(* IEC 61131-3 sources: programs/VI-54/VI-54_20171205/VI-54_20171205/Stations/PLC_VI54/VI-54_171014/Class/_DriveAxisBase (part 2) *)

  //Error of Axis gets only shown, if Axis is Online
  if bOnlineFinished then
    AxError := GetAxError();
  else
    AxError := 0;
  end_if;

  output := AxError;

END_FUNCTION

FUNCTION _DriveAxisBase::LoadDrivePara
  VAR
    pTabAdress : ^DINT;
    TabLength   : DINT;
  END_VAR

  // load the parameter data to the para objects
  case DriveInitType of

    _SDDSTDTABLE :

     pTabAdress := GetTabAdress(TabType:= 0, bdSettings.bSendMPara, #TabLength);
     SetListToParObj(pData:= (pTabAdress)$^DINT, udLen:=TabLength$UDINT);

    _SDDL2TABLE :
    // load the data of the table
      pTabAdress := GetTabAdress(TabType:= 1, bdSettings.bSendMPara, #TabLength);
      SetListToParObj(pData:= (pTabAdress)$^DINT, udLen:=TabLength$UDINT);

    _SDDRAMEX,
    _SDDFILE :
      pSDDData$^void := DriveAxisSet.GetMemPtr();
      if pSDDData <> NIL then
        // load the data of the memory
        SetListToParObj(pData:= (pSDDData$DINT + pSDDData^.AxOffset)$^DINT, udLen:=pSDDData^.AxLength);
      end_if;

  end_case;

END_FUNCTION

FUNCTION _DriveAxisBase::SetListToParObj
	VAR_INPUT
		pData 	: ^DINT;
		udLen 	: UDINT;
	END_VAR
	VAR_OUTPUT
		retcode 	: BOOL;
	END_VAR
  VAR
    pHlp          : ^DINT;
    x             : UDINT;
    pThisNewInst  : ^void;
    usParaNr      : USINT;
    ParaValue     : DINT;
    UserPara      : CmdStruct;
    UserResult    : Results;
  END_VAR

  retcode := FALSE;

  //hier konnte es zu einem Problem kommen kann wenn pThisNewInst nicht init war.
  pThisNewInst := NIL; //BleErn 19.08.2010 11:27

  if (bdSettings.bAxSetPara = FALSE) | (pData = NIL) then
    return;
  end_if;

  x := 0;
  pHlp := pData;

  while x < udLen do

    usParaNr := pHlp^$USINT;
    pHlp += sizeof(USINT);
    x += sizeof(USINT);

    if usParaNr <= MAX_MOTOR_PARA then
      pThisNewInst$DINT := AxSetPara[IDX_MOTOR_PARA];
    elsif usParaNr <= MAX_DRIVE_PARA then
      pThisNewInst$DINT := AxSetPara[IDX_DRIVE_PARA];
    elsif usParaNr <= MAX_CURRENT_PARA then
      pThisNewInst$DINT := AxSetPara[IDX_CURRENT_PARA];
    elsif usParaNr <= MAX_VEL_PARA then
      pThisNewInst$DINT := AxSetPara[IDX_VEL_PARA];
    elsif usParaNr <= MAX_POS_PARA then
      pThisNewInst$DINT := AxSetPara[IDX_POS_PARA];
    elsif usParaNr <= MAX_FD_PARA then
      pThisNewInst$DINT := AxSetPara[IDX_FD_PARA];
    elsif usParaNr <= MAX_APPLI_PARA then
      pThisNewInst$DINT := AxSetPara[IDX_APPLI_PARA];
    elsif usParaNr <= MAX_ERRORHANDLING then
      pThisNewInst$DINT := AxSetPara[IDX_ERRORHANDLING];
    end_if;

    ParaValue := pHlp^$DINT;
    if pThisNewInst <> NIL then
      UserPara.uiCmd := SDD_REFRESH_SETPARA;
      UserPara.aPara[0] := to_dint(usParaNr);
      UserPara.aPara[1] := ParaValue;
      pThisNewInst$^VirtualBase^.NewInst(#UserPara, #UserResult);
    end_if;

    pHlp += sizeof(UDINT);
    x += sizeof(UDINT);

  end_while;

END_FUNCTION

FUNCTION VIRTUAL GLOBAL _DriveAxisBase::SDDProcess

  //SA 23391 - ObeChr: Wait for Online before starting SDDCmdInterface
  if Online = 1 then

    case SDDCmdIntfc of

    _SDDIDLE :
      // do nothing

    _SDDREADALL :
      if bdSettings.bStartRead = FALSE then
        bdSettings.bStartRead := TRUE;
        // check if a read is possible
        if ChkParaRead(0) = FALSE then
          SDDCmdIntfc := _SDDIDLE;
        else
          ParaReadProc();
        end_if;
      else
        // überprüfen ob alle Parameter schon vorhanden sind
        ParaReadProc();
        if (bdSettings.bReadAxFin = TRUE) then
          SDDCmdIntfc := _SDDIDLE;
          bdSettings.bStartRead := FALSE;
        end_if;
      end_if;

    _SDDINIT :

      if (AxEnable = 0)  then
        if OldSDDCmdIntfc <> SDDCmdIntfc then
          DriveMng.InitDrive(0); // start the initialisation of the drive
          Init_Again:=true;
          //bdSettings.bDriveInitialized:=true;
        end_if;
      else
        SDDCmdIntfc := _SDDIDLE;
      end_if;

    _SDDURINIT :

      if (AxEnable = 0) then
        if OldSDDCmdIntfc <> SDDCmdIntfc then
          DriveMng.InitDrive(1); // start the initialisation of the drive
          InitASyncPara(); // initialize the structure
          Init_Again:=true;
        end_if;
      else
        SDDCmdIntfc := _SDDIDLE;
      end_if;

    _SDDEXDATA :

      // only if a object of the correct class is connected
      if DriveAxisSet.ChkFileHandle() then

        if OldSDDCmdIntfc <> SDDCmdIntfc then
          pSDDData$^void := DriveAxisSet.GetMemPtr();

          _strcpy(#pSDDData^.AxName[0],#szObjName[0]); //here the name of the object is set to the struct
          DriveAxisSet.SetUserSSDCmd(_SDDEXDATA, pSDDData);
        else
          SDDCmdIntfc := DriveAxisSet.GetUserSSDCmd();
        end_if;
      else
        SDDCmdIntfc := _SDDIDLE;
      end_if;

    end_case;

    OldSDDCmdIntfc := SDDCmdIntfc;

  end_if;

END_FUNCTION

FUNCTION VIRTUAL GLOBAL _DriveAxisBase::SDDCmdIntfc::Write
	VAR_INPUT
		input (EAX) 	: _SDDUSERCMD;
	END_VAR
	VAR_OUTPUT
		result (EAX) 	: _SDDUSERCMD;
	END_VAR

  if SDDCmdIntfc = _SDDIDLE then
    SDDCmdIntfc := input;
    result := SDDCmdIntfc;
  else
    result$DINT := ACCESS_DENIED;
  end_if;

END_FUNCTION

FUNCTION _DriveAxisBase::ChkParaRead
	VAR_INPUT
		ChkType 	: DINT;
	END_VAR
	VAR_OUTPUT
		retcode 	: BOOL;
	END_VAR

  retcode := FALSE;

  case ChkType of
  0 : // check if a reading command is allowed

    bdSettings.bReadAx := FALSE;

    bdSettings.bReadAxFin := FALSE;

    if (bdSettings.bAxSetPara = TRUE)then
      bdSettings.bReadAx := TRUE;
      ParaReadCmdAx := 1;
      retcode := TRUE;
    else
      bdSettings.bReadAxFin := TRUE;
    end_if;

  1 : // check if we can send the next reading commands
    if ParaReadCmdAx = 2 then
      if AxASyncPara.ActEntries < 10 then
        retcode := TRUE;
      end_if;
    end_if;

  end_case;

END_FUNCTION

FUNCTION _DriveAxisBase::ParaReadProc
  VAR
    dValue      : DINT;
    pThis       : ^void;
    i           : DINT;
    UserPara    : CmdStruct;
    UserResult  : Results;
  END_VAR
        // Start laden aller Parameter vom Drive
        // folgender Ablauf :
        // 1. Es wird für jede Achse die Anforderung in den Ringbuffer geschrieben (30mal).(Eigene Kennung erforderlich ?);
        // 2. Warten bis nur mehr 10 Einträge vorhanden sind, und dann die nächsten Einträge absetzen
        // 3. wenn alle Einträge abgesetzt sind, (letzter Eintrag muss eine extra Kennung haben), wird überprüft wann alle Daten vorhanden sind
        // 4. Wenn ein Wert eines Parameters ankommt, wird dieser in den Speicher geschrieben, dies ist abhängig von der Sicherungsauswahl. Ist eine Tabelle ausgewählt
        //    werden die Daten sofort an die Parameterklassen gesendet, sind keine Parameterobjekte vorhanden, so wird der Vorgang gar nicht durchgeführt.
        // 5. Wenn der letzte Wert des Parameters kommt, wird die Chksumme neu berechnet, die Daten weggesichert, und die Parameterobjekte aktualisiert

  dValue := 0;

 if bdSettings.bReadAx = TRUE then
    case ParaReadCmdAx of

    0 : //idle step

    1 : // set the first entries in the buffer
      // set the info busy to all para classes
      UserPara.uiCmd := SDD_ASYNC_BUSY;

      for i := IDX_MOTOR_PARA to IDX_ERRORHANDLING do
        pThis$DINT := AxSetPara[i];
        if pThis <> NIL then
          // Set the state BUSY
          pThis$^VirtualBase^.NewInst(#UserPara, #UserResult);
        end_if;
      end_for;

      if AxSetPara[IDX_MOTOR_PARA] <> 0 then
        pThis$DINT := AxSetPara[IDX_MOTOR_PARA];

        AddASyncEntry(usParaNr:= SDD_M_NAME1, usRdWr:= 0, dValue:= dValue, pThisObj:= pThis, usEntry:= 1);
        AddASyncEntry(usParaNr:= SDD_M_NAME2, usRdWr:= 0, dValue:= dValue, pThisObj:= pThis, usEntry:= 1);
        AddASyncEntry(usParaNr:= SDD_M_NAME3, usRdWr:= 0, dValue:= dValue, pThisObj:= pThis, usEntry:= 1);
        AddASyncEntry(usParaNr:= SDD_M_INULL, usRdWr:= 0, dValue:= dValue, pThisObj:= pThis, usEntry:= 1);
        AddASyncEntry(usParaNr:= SDD_M_IPEAK, usRdWr:= 0, dValue:= dValue, pThisObj:= pThis, usEntry:= 1);
        AddASyncEntry(usParaNr:= SDD_M_NMAX, usRdWr:= 0, dValue:= dValue, pThisObj:= pThis, usEntry:= 1);
        AddASyncEntry(usParaNr:= SDD_M_POL, usRdWr:= 0, dValue:= dValue, pThisObj:= pThis, usEntry:= 1);
        AddASyncEntry(usParaNr:= SDD_M_TORQUE, usRdWr:= 0, dValue:= dValue, pThisObj:= pThis, usEntry:= 1);
        AddASyncEntry(usParaNr:= SDD_M_L, usRdWr:= 0, dValue:= dValue, pThisObj:= pThis, usEntry:= 1);
        AddASyncEntry(usParaNr:= SDD_M_R, usRdWr:= 0, dValue:= dValue, pThisObj:= pThis, usEntry:= 1);
        AddASyncEntry(usParaNr:= SDD_M_J, usRdWr:= 0, dValue:= dValue, pThisObj:= pThis, usEntry:= 1);
        AddASyncEntry(usParaNr:= SDD_M_TYPE, usRdWr:= 0, dValue:= dValue, pThisObj:= pThis, usEntry:= 1);
        AddASyncEntry(usParaNr:= SDD_M_RPOL, usRdWr:= 0, dValue:= dValue, pThisObj:= pThis, usEntry:= 1);
        AddASyncEntry(usParaNr:= SDD_M_ROFF, usRdWr:= 0, dValue:= dValue, pThisObj:= pThis, usEntry:= 1);
        AddASyncEntry(usParaNr:= SDD_M_RPULSE, usRdWr:= 0, dValue:= dValue, pThisObj:= pThis, usEntry:= 1);
        AddASyncEntry(usParaNr:= SDD_M_RTEMP, usRdWr:= 0, dValue:= dValue, pThisObj:= pThis, usEntry:= 1);
        AddASyncEntry(usParaNr:= SDD_M_SER, usRdWr:= 0, dValue:= dValue, pThisObj:= pThis, usEntry:= 1);
        AddASyncEntry(usParaNr:= SDD_M_BRAKE, usRdWr:= 0, dValue:= dValue, pThisObj:= pThis, usEntry:= 1);
        AddASyncEntry(usParaNr:= SDD_M_IFWEAK, usRdWr:= 0, dValue:= dValue, pThisObj:= pThis, usEntry:= 1);
        AddASyncEntry(usParaNr:= SDD_M_BRDIS, usRdWr:= 0, dValue:= dValue, pThisObj:= pThis, usEntry:= 1);
        AddASyncEntry(usParaNr:= SDD_M_BREN, usRdWr:= 0, dValue:= dValue, pThisObj:= pThis, usEntry:= 1);
        AddASyncEntry(usParaNr:= SDD_M_IMAG, usRdWr:= 0, dValue:= dValue, pThisObj:= pThis, usEntry:= 1);
        AddASyncEntry(usParaNr:= SDD_M_TROT, usRdWr:= 0, dValue:= dValue, pThisObj:= pThis, usEntry:= 1);
        AddASyncEntry(usParaNr:= SDD_M_UN, usRdWr:= 0, dValue:= dValue, pThisObj:= pThis, usEntry:= 1);
        AddASyncEntry(usParaNr:= SDD_M_UBOOST, usRdWr:= 0, dValue:= dValue, pThisObj:= pThis, usEntry:= 1);
      end_if;

      if AxSetPara[IDX_DRIVE_PARA] <> 0 then
        pThis$DINT := AxSetPara[IDX_DRIVE_PARA];
        AddASyncEntry(usParaNr:= SDD_G_MODE, usRdWr:= 0, dValue:= dValue, pThisObj:= pThis, usEntry:= 1);
        AddASyncEntry(usParaNr:= SDD_G_CETIME, usRdWr:= 0, dValue:= dValue, pThisObj:= pThis, usEntry:= 1);
        AddASyncEntry(usParaNr:= SDD_G_VMAINS, usRdWr:= 0, dValue:= dValue, pThisObj:= pThis, usEntry:= 1);
        AddASyncEntry(usParaNr:= SDD_G_VBUSM, usRdWr:= 0, dValue:= dValue, pThisObj:= pThis, usEntry:= 1);
        AddASyncEntry(usParaNr:= SDD_G_VBUSM, usRdWr:= 0, dValue:= dValue, pThisObj:= pThis, usEntry:= 1);
        AddASyncEntry(usParaNr:= SDD_G_MTEMPK, usRdWr:= 0, dValue:= dValue, pThisObj:= pThis, usEntry:= 1);
        AddASyncEntry(usParaNr:= SDD_G_MTEMPE, usRdWr:= 0, dValue:= dValue, pThisObj:= pThis, usEntry:= 1);
        AddASyncEntry(usParaNr:= SDD_G_PWM, usRdWr:= 0, dValue:= dValue, pThisObj:= pThis, usEntry:= 1);
        AddASyncEntry(usParaNr:= SDD_G_DELAY, usRdWr:= 0, dValue:= dValue, pThisObj:= pThis, usEntry:= 1);
        AddASyncEntry(usParaNr:= SDD_G_FTEMP, usRdWr:= 0, dValue:= dValue, pThisObj:= pThis, usEntry:= 1);
        AddASyncEntry(usParaNr:= SDD_G_EMRAMP, usRdWr:= 0, dValue:= dValue, pThisObj:= pThis, usEntry:= 1);
        AddASyncEntry(usParaNr:= SDD_G_MASKE1, usRdWr:= 0, dValue:= dValue, pThisObj:= pThis, usEntry:= 1);
        AddASyncEntry(usParaNr:= SDD_G_MASKE2, usRdWr:= 0, dValue:= dValue, pThisObj:= pThis, usEntry:= 1);
        AddASyncEntry(usParaNr:= SDD_G_MASKW, usRdWr:= 0, dValue:= dValue, pThisObj:= pThis, usEntry:= 1);
        AddASyncEntry(usParaNr:= SDD_G_MASKD, usRdWr:= 0, dValue:= dValue, pThisObj:= pThis, usEntry:= 1);
        AddASyncEntry(usParaNr:= SDD_G_VRAMP, usRdWr:= 0, dValue:= dValue, pThisObj:= pThis, usEntry:= 1);
        AddASyncEntry(usParaNr:= SDD_G_SRAMP, usRdWr:= 0, dValue:= dValue, pThisObj:= pThis, usEntry:= 1);
        AddASyncEntry(usParaNr:= SDD_G_RBAL, usRdWr:= 0, dValue:= dValue, pThisObj:= pThis, usEntry:= 1);
      end_if;

      ParaReadCmdAx := 2;

    2 :
      // wait until only 10 entries in the buffer

      if ChkParaRead(ChkType:= 1) = TRUE then
        ParaReadCmdAx := 3;
      end_if;

    3 :
      // send the rest

      if AxSetPara[IDX_CURRENT_PARA] <> 0 then
        pThis$DINT := AxSetPara[IDX_CURRENT_PARA];
        AddASyncEntry(usParaNr:= SDD_C_KPQ, usRdWr:= 0, dValue:= dValue, pThisObj:= pThis, usEntry:= 1);
        AddASyncEntry(usParaNr:= SDD_C_TN, usRdWr:= 0, dValue:= dValue, pThisObj:= pThis, usEntry:= 1);
        AddASyncEntry(usParaNr:= SDD_C_KDREL, usRdWr:= 0, dValue:= dValue, pThisObj:= pThis, usEntry:= 1);
        AddASyncEntry(usParaNr:= SDD_C_KPDREL, usRdWr:= 0, dValue:= dValue, pThisObj:= pThis, usEntry:= 1);
        AddASyncEntry(usParaNr:= SDD_C_KPNULL, usRdWr:= 0, dValue:= dValue, pThisObj:= pThis, usEntry:= 1);
        AddASyncEntry(usParaNr:= SDD_C_KPPEAK, usRdWr:= 0, dValue:= dValue, pThisObj:= pThis, usEntry:= 1);
        AddASyncEntry(usParaNr:= SDD_C_ICONT, usRdWr:= 0, dValue:= dValue, pThisObj:= pThis, usEntry:= 1);
        AddASyncEntry(usParaNr:= SDD_C_IPEAK, usRdWr:= 0, dValue:= dValue, pThisObj:= pThis, usEntry:= 1);
        AddASyncEntry(usParaNr:= SDD_C_IPEAKN, usRdWr:= 0, dValue:= dValue, pThisObj:= pThis, usEntry:= 1);
      end_if;

      if AxSetPara[IDX_VEL_PARA] <> 0 then
        pThis$DINT := AxSetPara[IDX_VEL_PARA];
        AddASyncEntry(usParaNr:= SDD_V_KP, usRdWr:= 0, dValue:= dValue, pThisObj:= pThis, usEntry:= 1);
        AddASyncEntry(usParaNr:= SDD_V_TN, usRdWr:= 0, dValue:= dValue, pThisObj:= pThis, usEntry:= 1);
        AddASyncEntry(usParaNr:= SDD_V_T, usRdWr:= 0, dValue:= dValue, pThisObj:= pThis, usEntry:= 1);
        AddASyncEntry(usParaNr:= SDD_V_T2, usRdWr:= 0, dValue:= dValue, pThisObj:= pThis, usEntry:= 1);
        AddASyncEntry(usParaNr:= SDD_V_FILT, usRdWr:= 0, dValue:= dValue, pThisObj:= pThis, usEntry:= 1);
        AddASyncEntry(usParaNr:= SDD_V_NMAX, usRdWr:= 0, dValue:= dValue, pThisObj:= pThis, usEntry:= 1);
        AddASyncEntry(usParaNr:= SDD_V_KPREL, usRdWr:= 0, dValue:= dValue, pThisObj:= pThis, usEntry:= 1);
      end_if;

      if AxSetPara[IDX_POS_PARA] <> 0 then
        pThis$DINT := AxSetPara[IDX_POS_PARA];
        AddASyncEntry(usParaNr:= SDD_P_KV, usRdWr:= 0, dValue:= dValue, pThisObj:= pThis, usEntry:= 1);
        AddASyncEntry(usParaNr:= SDD_P_SFF, usRdWr:= 0, dValue:= dValue, pThisObj:= pThis, usEntry:= 1);
        AddASyncEntry(usParaNr:= SDD_P_PSCALE, usRdWr:= 0, dValue:= dValue, pThisObj:= pThis, usEntry:= 1);
        AddASyncEntry(usParaNr:= SDD_P_SSCALE, usRdWr:= 0, dValue:= dValue, pThisObj:= pThis, usEntry:= 1);
        AddASyncEntry(usParaNr:= SDD_P_TFF, usRdWr:= 0, dValue:= dValue, pThisObj:= pThis, usEntry:= 1);
        AddASyncEntry(usParaNr:= SDD_P_PEMAX, usRdWr:= 0, dValue:= dValue, pThisObj:= pThis, usEntry:= 1);
        AddASyncEntry(usParaNr:= SDD_P_SMODE, usRdWr:= 0, dValue:= dValue, pThisObj:= pThis, usEntry:= 1);
      end_if;

      if AxSetPara[IDX_FD_PARA] <> 0 then
        pThis$DINT := AxSetPara[IDX_FD_PARA];
        AddASyncEntry(usParaNr:= SDD_F_BW, usRdWr:= 0, dValue:= dValue, pThisObj:= pThis, usEntry:= 1);
        AddASyncEntry(usParaNr:= SDD_F_FF, usRdWr:= 0, dValue:= dValue, pThisObj:= pThis, usEntry:= 1);
        AddASyncEntry(usParaNr:= SDD_F_RK, usRdWr:= 0, dValue:= dValue, pThisObj:= pThis, usEntry:= 1);
      end_if;

      if AxSetPara[IDX_APPLI_PARA] <> 0 then
        pThis$DINT := AxSetPara[IDX_APPLI_PARA];
        AddASyncEntry(usParaNr:= SDD_A_JRATIO, usRdWr:= 0, dValue:= dValue, pThisObj:= pThis, usEntry:= 1);
        AddASyncEntry(usParaNr:= SDD_A_VALRT1, usRdWr:= 0, dValue:= dValue, pThisObj:= pThis, usEntry:= 1);
        AddASyncEntry(usParaNr:= SDD_A_VALRT2, usRdWr:= 0, dValue:= dValue, pThisObj:= pThis, usEntry:= 1);
        AddASyncEntry(usParaNr:= SDD_A_VALTT1, usRdWr:= 0, dValue:= dValue, pThisObj:= pThis, usEntry:= 1);
        AddASyncEntry(usParaNr:= SDD_A_VALTT2, usRdWr:= 0, dValue:= dValue, pThisObj:= pThis, usEntry:= 1);
        AddASyncEntry(usParaNr:= SDD_A_CTIME, usRdWr:= 0, dValue:= dValue, pThisObj:= pThis, usEntry:= 1);
        AddASyncEntry(usParaNr:= SDD_A_STIME, usRdWr:= 0, dValue:= dValue, pThisObj:= pThis, usEntry:= 1);
        AddASyncEntry(usParaNr:= SDD_A_STYPE, usRdWr:= 0, dValue:= dValue, pThisObj:= pThis, usEntry:= 1);
        AddASyncEntry(usParaNr:= SDD_A_AVSW, usRdWr:= 0, dValue:= dValue, pThisObj:= pThis, usEntry:= 1);
        AddASyncEntry(usParaNr:= SDD_A_I2TERR, usRdWr:= 0, dValue:= dValue, pThisObj:= pThis, usEntry:= 1);
        AddASyncEntry(usParaNr:= SDD_A_TEMPDE, usRdWr:= 0, dValue:= dValue, pThisObj:= pThis, usEntry:= 1);
        AddASyncEntry(usParaNr:= SDD_A_TEMPMW, usRdWr:= 0, dValue:= dValue, pThisObj:= pThis, usEntry:= 1);
        AddASyncEntry(usParaNr:= SDD_A_STRED, usRdWr:= 0, dValue:= dValue, pThisObj:= pThis, usEntry:= 1);
        AddASyncEntry(usParaNr:= SDD_A_STDT, usRdWr:= 0, dValue:= dValue, pThisObj:= pThis, usEntry:= 1);
        AddASyncEntry(usParaNr:= SDD_A_POS, usRdWr:= 0, dValue:= dValue, pThisObj:= pThis, usEntry:= 1);
        AddASyncEntry(usParaNr:= SDD_A_DNAME1, usRdWr:= 0, dValue:= dValue, pThisObj:= pThis, usEntry:= 1);
        AddASyncEntry(usParaNr:= SDD_A_DNAME2, usRdWr:= 0, dValue:= dValue, pThisObj:= pThis, usEntry:= 1);
        AddASyncEntry(usParaNr:= SDD_A_DNAME3, usRdWr:= 0, dValue:= dValue, pThisObj:= pThis, usEntry:= 1);
        AddASyncEntry(usParaNr:= SDD_A_MODE2, usRdWr:= 0, dValue:= dValue, pThisObj:= pThis, usEntry:= 1);
        AddASyncEntry(usParaNr:= SDD_A_MULTI, usRdWr:= 0, dValue:= dValue, pThisObj:= pThis, usEntry:= 1);
        AddASyncEntry(usParaNr:= SDD_A_CAPREF, usRdWr:= 0, dValue:= dValue, pThisObj:= pThis, usEntry:= 1);
        AddASyncEntry(usParaNr:= SDD_A_EDGE, usRdWr:= 0, dValue:= dValue, pThisObj:= pThis, usEntry:= 1);
        AddASyncEntry(usParaNr:= SDD_A_STTH, usRdWr:= 0, dValue:= dValue, pThisObj:= pThis, usEntry:= 1);
        AddASyncEntry(usParaNr:= SDD_A_INT1, usRdWr:= 0, dValue:= dValue, pThisObj:= pThis, usEntry:= 1);
        AddASyncEntry(usParaNr:= SDD_A_INT2, usRdWr:= 0, dValue:= dValue, pThisObj:= pThis, usEntry:= 1);
        AddASyncEntry(usParaNr:= SDD_A_ICOM, usRdWr:= 0, dValue:= dValue, pThisObj:= pThis, usEntry:= 1);
        AddASyncEntry(usParaNr:= SDD_A_ICOMP, usRdWr:= 0, dValue:= dValue, pThisObj:= pThis, usEntry:= 1);
        AddASyncEntry(usParaNr:= SDD_A_CMIN, usRdWr:= 0, dValue:= dValue, pThisObj:= pThis, usEntry:= 1);
        AddASyncEntry(usParaNr:= SDD_A_BIQCF, usRdWr:= 0, dValue:= dValue, pThisObj:= pThis, usEntry:= 1);
        AddASyncEntry(usParaNr:= SDD_A_BIQFR, usRdWr:= 0, dValue:= dValue, pThisObj:= pThis, usEntry:= 1);
        AddASyncEntry(usParaNr:= SDD_A_BIQCD, usRdWr:= 0, dValue:= dValue, pThisObj:= pThis, usEntry:= 1);
        AddASyncEntry(usParaNr:= SDD_A_BIQDR, usRdWr:= 0, dValue:= dValue, pThisObj:= pThis, usEntry:= 1);
        AddASyncEntry(usParaNr:= SDD_A_CAPFT, usRdWr:= 0, dValue:= dValue, pThisObj:= pThis, usEntry:= 1);
      end_if;

      if AxSetPara[IDX_ERRORHANDLING] <> 0 then
        pThis$DINT := AxSetPara[IDX_ERRORHANDLING];
        AddASyncEntry(usParaNr:= SDD_I_STATUS, usRdWr:= 0, dValue:= dValue, pThisObj:= pThis, usEntry:= 1);
        AddASyncEntry(usParaNr:= SDD_I_DERROR, usRdWr:= 0, dValue:= dValue, pThisObj:= pThis, usEntry:= 1);
      end_if;

      // get the number of parameters in the drive (only to know if we are at the end of the reading process
      AddASyncEntry(usParaNr:= 0, usRdWr:= 0, dValue:= dValue, pThisObj:= NIL, usEntry:= 2);
      ParaReadCmdAx := 4;
    4 :

      if bdSettings.bReadAxFin = TRUE then
      // wait until the last entry is send the value back

        // now save all parameters in the SRAM / FILE
        if DriveInitType = _SDDRAMEX then
          pSDDData$^void := DriveAxisSet.GetMemPtr();
          DriveAxisSet.SaveRamExData(pData:= pSDDData, udLen:= pSDDData^.udLen, udOffset:= 0);

        elsif DriveInitType = _SDDFILE then
          pSDDData$^void := DriveAxisSet.GetMemPtr();
          DriveAxisSet.SaveRamFileData(pData:= pSDDData, udLen:= pSDDData^.udLen, udOffset:= 0);

        end_if;
        ParaReadCmdAx := 0;

      end_if;
    end_case;
  end_if;

END_FUNCTION

FUNCTION VIRTUAL GLOBAL _DriveAxisBase::SetAbsolutePosition
	VAR_INPUT
		AbsPosition 	: DINT;
	END_VAR
	VAR_OUTPUT
		retcode 	: DINT;
	END_VAR

  retcode := 1;
  if IsOnline() = FALSE then
    retcode := -1;  // no communication available or the initialisation isn't finished
    return;
  end_if;

  //Check if operation is already in progress
  if bdSettings.bSetAbsPos = true then
    retcode := -2;
    return;
  end_if;

  // check if the axis is with an absolute encoder
  if (bdSettings.bNoAbsEnc = FALSE) then
    // if any axis is enabled, the parameter K-FBRW cannot be written
    if DriveMng.IsAnyAxisEnabled() then
      retcode := -4;
      return;
    end_if;

    // set the value of the parameter A-MULTI to 1
    AddASyncEntry(SDD_A_MULTI, 1, 1, this, 0);
    // set the new position to the parameter
    AddASyncEntry(SDD_A_POS, 1, AbsPosition, this, 1);
    // marry the motor with the Drive
    AddASyncEntry(SDD_K_FBRW, 1, 3, this, 1);

    bdSettings.bSetAbsPos := TRUE;
  else
    retcode := -3; // no absolute encoder available
  end_if;

END_FUNCTION

FUNCTION VIRTUAL GLOBAL _DriveAxisBase::SetAbsolutePositionEncoder
	VAR_INPUT
		AbsPosition 	: DINT;
	END_VAR
	VAR_OUTPUT
		retcode 	: DINT;
	END_VAR

  //Init Returncode
  retcode := true;

  //Check if Drive is Online and the Initialization is finished
  if IsOnline() = false then
    retcode := -1;
    return;
  end_if;

  //Check if operation is already in progress
  if bdSettings.bSetAbsPosEncoder = true then
    retcode := -2;
    return;
  end_if;

  //Check if the Axis got an AbsoluteEncoder
  if bdSettings.bNoAbsEnc = false then
    // if axis is enabled, the parameter K-FBRW cannot be written
    if DriveMng.IsAnyAxisEnabled() then
      retcode := -4;
      return;
    end_if;

    //Set A-MULTI to 1
    AddASyncEntry(SDD_A_MULTI, true, 0, this, 0);

    //Set A-POS to InputParamter
    AddASyncEntry(SDD_A_POS, true, AbsPosition, this, 1);

    //Set K-FBRW to 5 => Calculate Offset
    AddASyncEntry(SDD_K_FBRW, true, 5, this, 1);

    //Set K-FBRW to 2 => Save Offset in Feedback
    AddASyncEntry(SDD_K_FBRW, true, 2, this, 1);

    bdSettings.bSetAbsPosEncoder := true;
  else
    retcode := -3;
  end_if;

END_FUNCTION

FUNCTION _DriveAxisBase::SaveDrivePara
  VAR
    TabAddress 	: ^DINT;
    pHlpSDD		: ^void;
    TabLength   : DINT;
  END_VAR

  // get the actual ptr of the memory
  pSDDData$^void := DriveAxisSet.GetMemPtr();

  if pSDDData <> NIL then

    pSDDData^.udLen := sizeof(_SDDMEMHEADER); // initialize the length of the data
    pSDDData^.AxOffset := sizeof(_SDDMEMHEADER); // set the offset
    TabAddress := GetTabAdress(1, bdSettings.bSendMPara, #TabLength);

    if TabAddress = NIL then
      return;
    end_if;

    pSDDData^.AxLength := TabLength$UDINT;

    pHlpSDD := pSDDData + pSDDData^.AxOffset;

    _memcpy(pHlpSDD, (TabAddress)$^void, (TabLength)$UDINT);

    pSDDData^.udLen += pSDDData^.AxLength;

    // calculate the crc of the sdd parameters
    pSDDData^.udCRC32 := CalcCRC32((pSDDData + sizeof(UDINT))$^UDINT, pSDDData^.udLen - sizeof(UDINT));

    case DriveInitType of

    _SDDRAMEX :

      // save the data in the ramex
      DriveAxisSet.SaveRamExData(pSDDData, pSDDData^.udLen, 0);

    _SDDFILE :
      // save the data in the ramfile
      DriveAxisSet.SaveRamFileData(pSDDData, pSDDData^.udLen, 0);

    end_case;
  end_if;

END_FUNCTION

FUNCTION _DriveAxisBase::CalcCRC32
	VAR_INPUT
		pData 	: ^UDINT;
		udLen 	: UDINT;
	END_VAR
	VAR_OUTPUT
		CRC32 	: UDINT;
	END_VAR

	CRC32 := coLinker.CRC32(0, pData$^void, udLen);

END_FUNCTION

FUNCTION VIRTUAL GLOBAL _DriveAxisBase::GetZImpulse
	VAR_OUTPUT
		retcode 	: USINT;
	END_VAR

  retcode:=0;

  if ( ( ActPos and maskZImpulse$DINT ) <> oldRevolutions ) then
    retcode := 1;
    oldRevolutions := (ActPos and maskZImpulse$DINT);
  end_if;

END_FUNCTION

FUNCTION VIRTUAL GLOBAL _DriveAxisBase::ZPulsLatch::Read
	VAR_OUTPUT
		output (EAX) 	: DINT;
	END_VAR

  if bOnlineFinished then

    if ZPulsLatch = 0 then
      output := ZPulsLatch := GetZImpulse();
    else
      output := ZPulsLatch;
      ZPulsLatch := 0;
    end_if;

  else
    ZPulsLatch := 0;
    output := ZPulsLatch;
  end_if;

END_FUNCTION

FUNCTION _DriveAxisBase::SetZPulseMask

  maskZImpulse:=16#FFFFFFFF;
  maskZImpulse:=maskZImpulse SHL (32-ppscale);

  //P-PSCALE  0: 00000000 00000000 00000000 00000000
  //P-PSCALE 10: 11111111 11000000 00000000 00000000
  //P-PSCALE 16: 11111111 11111111 00000000 00000000

END_FUNCTION

FUNCTION VIRTUAL GLOBAL _DriveAxisBase::GetSyncEntry
	VAR_INPUT
		usValue 	: USINT;
		usPData 	: ^DINT;
	END_VAR
	VAR_OUTPUT
		retcode 	: DINT;
	END_VAR

  retcode:=DriveMng.GetSyncEntry(usAxis:=usAxisIndex, usValue:=usValue, usPData:=usPData);

END_FUNCTION

FUNCTION VIRTUAL GLOBAL _DriveAxisBase::AddSyncEntry
	VAR_INPUT
		pThis 	: ^void;
	END_VAR
	VAR_OUTPUT
		retcode 	: BOOL;
	END_VAR

  retcode := FALSE;

  if pThis <> NIL then
    SyncParaObject := pThis$DINT;
    retcode := TRUE;
  end_if;

END_FUNCTION

FUNCTION VIRTUAL GLOBAL _DriveAxisBase::SetSyncEntry
	VAR_INPUT
		usValue 	: USINT;
		usPData 	: DINT;
	END_VAR
	VAR_OUTPUT
		retcode 	: DINT;
	END_VAR

  retcode:=DriveMng.SetSyncEntry(usAxis:=usAxisIndex, usValue:=usValue, usPData:=usPData);

END_FUNCTION

FUNCTION _DriveAxisBase::RefreshIASP
	VAR_INPUT
		Para 	  : DINT;
		Value 	: DINT;
	END_VAR
  VAR
  	UserPara      : CmdStruct;
    UserResult    : Results;
  END_VAR

  // if there is a change in the following values, first we set the pointers to zero, and then we initialize them, allready with the new value

  if AxEnable = 0 then //just do some changes when the axis does not run
    case Para of
      SDD_A_VALTT1:

        _memset(#SyncPara.ActCurrent,0,sizeof(SyncPara.ActCurrent));
        _memset(#SyncPara.ActPos,    0,sizeof(SyncPara.ActPos));
        _memset(#SyncPara.ActSpeed,  0,sizeof(SyncPara.ActSpeed));
        _memset(#SyncPara.Xw,        0,sizeof(SyncPara.Xw));
        _memset(#SyncPara.StateWord, 0,sizeof(SyncPara.StateWord));

        ActValues[0] := to_usint( Value AND 16#000000FF);
        ActValues[1] := to_usint((Value AND 16#0000FF00) SHR 8);

        GetSynchronPara();

      SDD_A_VALTT2:

        _memset(#SyncPara.ActCurrent,0,sizeof(SyncPara.ActCurrent));
        _memset(#SyncPara.ActPos,    0,sizeof(SyncPara.ActPos));
        _memset(#SyncPara.ActSpeed,  0,sizeof(SyncPara.ActSpeed));
        _memset(#SyncPara.Xw,        0,sizeof(SyncPara.Xw));
        _memset(#SyncPara.StateWord, 0,sizeof(SyncPara.StateWord));

        ActValues[2] := to_usint( Value AND 16#000000FF);
        ActValues[3] := to_usint((Value AND 16#0000FF00) SHR 8);
        ActValues[4] := to_usint((Value AND 16#00FF0000) SHR 16);

        if (AxisExtend = 1) & (SyncParaObject<>NIL) then
          UserPara.uiCmd := 10;
          UserPara.aPara[2]:=ActValues[2];
          UserPara.aPara[3]:=ActValues[3];
          UserPara.aPara[4]:=ActValues[4];
          SyncParaObject$^VirtualBase^.pSvrChCmd.NewInst(#UserPara, #UserResult); //initialize also the extend class
        end_if;

        GetSynchronPara();

      SDD_A_VALRT1:

        _memset(#SyncPara.SetCurrent, 0,sizeof(SyncPara.SetCurrent));
        _memset(#SyncPara.SetPos,     0,sizeof(SyncPara.SetPos));
        _memset(#SyncPara.SetSpeed,   0,sizeof(SyncPara.SetSpeed));
        _memset(#SyncPara.SetTorque,  0,sizeof(SyncPara.SetTorque));
        _memset(#SyncPara.ControlWord,0,sizeof(SyncPara.ControlWord));

        SetValues[0] := to_usint( Value AND 16#000000FF);
        SetValues[1] := to_usint((Value AND 16#0000FF00) SHR 8);

        SetSynchronPara();
//        AxTorqueControl.Write(4500); //it does not matter which controlword we have, because the internal function reduced this amount to the top limit
        SetAxTorque(4500);

      SDD_A_VALRT2:

        _memset(#SyncPara.SetCurrent, 0,sizeof(SyncPara.SetCurrent));
        _memset(#SyncPara.SetPos,     0,sizeof(SyncPara.SetPos));
        _memset(#SyncPara.SetSpeed,   0,sizeof(SyncPara.SetSpeed));
        _memset(#SyncPara.SetTorque,  0,sizeof(SyncPara.SetTorque));
        _memset(#SyncPara.ControlWord,0,sizeof(SyncPara.ControlWord));

        SetValues[2] := to_usint( Value AND 16#000000FF);
        SetValues[3] := to_usint((Value AND 16#0000FF00) SHR 8);
        SetValues[4] := to_usint((Value AND 16#00FF0000) SHR 16);

        if (AxisExtend = 1) & (SyncParaObject<>NIL) then
          UserPara.uiCmd := 11;
          UserPara.aPara[2]:=SetValues[2];
          UserPara.aPara[3]:=SetValues[3];
          UserPara.aPara[4]:=SetValues[4];
          SyncParaObject$^VirtualBase^.pSvrChCmd.NewInst(#UserPara, #UserResult); //if there is a extend class connected, we have to initialize it
        end_if;

        SetSynchronPara();
//        AxTorqueControl.Write(4500); //it does not matter which controlword we have, because the internal function reduced this amount to the top limit
        SetAxTorque(4500);

      SDD_P_PSCALE:
        ppscale:=to_usint(Value);
        SetZPulseMask();

    end_case;
  end_if;

END_FUNCTION

FUNCTION VIRTUAL GLOBAL _DriveAxisBase::AxOkay
	VAR_OUTPUT
		retcode 	: DINT;
	END_VAR

  retcode := false;
  if AxisState = 0 then
    retcode := true;
  end_if;

END_FUNCTION

FUNCTION VIRTUAL GLOBAL _DriveAxisBase::Online::Read
	VAR_OUTPUT
		output (EAX) 	: DINT;
	END_VAR

  //--- if DriveMng is online, we have no internal error, and the error-reset after startup is ready, we say Online = 1
  Online := bOnlineFinished;

  output := Online;

END_FUNCTION

FUNCTION VIRTUAL GLOBAL _DriveAxisBase::ErrorQuitHandling
	VAR_INPUT
		input 	: DINT;
	END_VAR
	VAR_OUTPUT
		result 	: DINT;
	END_VAR

  AxErrorQuit:=input AND 1;

  // check if there is a control word mapped, before accessing the data
  if SyncPara.ControlWord.ptr then
    if (SyncPara.ControlWord.userinfo=0) then
      SyncPara.ControlWord.ptr^$BINT.2:=AxErrorQuit$BOOL; //FAULT RESET
    elsif(SyncPara.ControlWord.userinfo=1) then
      SyncPara.ControlWord.ptr^$BINT.8:=AxErrorQuit$BOOL; //FAULT RESET
    end_if;
  end_if;

  if AxErrorQuit = 1 then
    FirstErrorReset := 4;
    ErrorQuitTime:=ops.tAbsolute;
  end_if;

  Controlword.ResetFault := AxErrorQuit$BOOL;

  result := AxErrorQuit;

END_FUNCTION

FUNCTION VIRTUAL _DriveAxisBase::GetAxError
	VAR_OUTPUT
		AxError 	: DINT;
	END_VAR
  VAR
  	sBuffer      : BDINT; //StateWord Buffer
  END_VAR

  if SyncPara.StateWord.ptr<>NIL  then
    sBuffer := SyncPara.StateWord.ptr^$BDINT;
    AxError:=sBuffer.4; //the error is at both control words on the same place
  else
    AxError:=0;
  end_if;

END_FUNCTION

FUNCTION _DriveAxisBase::SetAxTorque
	VAR_INPUT
		NewTorque 	: UDINT;
	END_VAR
  VAR
    cBuffer       : BDINT; //ControlWord Buffer
  END_VAR

  // if we have a 16-Bit Controlword
  if SyncPara.SetTorque.userinfo = 0 then

    if NewTorque < 0 then
      NewTorque := 0;
    end_if;

    if NewTorque > 1000 then
      NewTorque := 1000;
    end_if;

    AxTorqueControl := NewTorque;

    //Check if pointer is valid
    if SyncPara.ControlWord.ptr then
      cBuffer:=SyncPara.ControlWord.ptr^$BDINT;
      SyncPara.SetTorque.ptr^$INT:= to_int(TorqueCalculation(cBuffer,NewTorque));
    end_if;

  elsif SyncPara.SetTorque.userinfo=1 then //that is for the 32-Bit Controlword

    if NewTorque < 0 then
      NewTorque := 0;
    end_if;

    if NewTorque > 4500 then
      NewTorque := 4500;
    end_if;

    AxTorqueControl := NewTorque;

    if SyncPara.SetTorque.ptr then
      SyncPara.SetTorque.ptr^$INT:=to_int(NewTorque);
    end_if;

  end_if;

END_FUNCTION

FUNCTION _DriveAxisBase::IsOnlineFinished
	VAR_OUTPUT
		bOnline 	: BOOL;
	END_VAR

  if (IsOnline() = TRUE) & (CmdState <> ERROR) & ((FirstErrorReset = 0) | (FirstErrorReset >= 4)) then
    bOnline := 1;
  else
    bOnline := 0;
  end_if;

END_FUNCTION

FUNCTION VIRTUAL GLOBAL _DriveAxisBase::AddASyncEntryDS402
	VAR_INPUT
		uiParaID 	  : UINT;
		usParaSubID : USINT;
		usRdWr 	    : USINT;
		pValue 	    : ^USINT;
		bsDataInfo 	: BSINT;
		pThisObj 	  : ^void;
		usEntry 	  : USINT;
	END_VAR
	VAR_OUTPUT
		retcode 	  : DINT;
	END_VAR

  retcode := DriveMng.AddASyncEntryDS402(AxisNo     := usAxisIndex
                                      , uiParaID    := uiParaID
                                      , usParaSubID := usParaSubID
                                      , usRdWr      := usRdWr
                                      , pValue      := pValue
                                      , bsDataInfo  := bsDataInfo
                                      , pThisObj    := pThisObj
                                      , usEntry     := usEntry
                                      );

END_FUNCTION
